// TIA Portal V19 export
FUNCTION_BLOCK "TIMER"   // FB5, LAD
{ S7_Optimized_Access := 'TRUE' }
// stored: MemoryReserve 100, SetENOAutomatically false
   VAR_INPUT
      START_TIMER : Bool;
      HR_SET : Int;
      MIN_SET : Int;
      SEC_SET : Int;
      RESET_TIMER : Bool;
   END_VAR
   VAR_OUTPUT
      SEC : Int;
      MIN : Int;
      HR : Int;
      TIMER_DONE { ExternalAccessible := 'False'; ExternalVisible := 'False'; ExternalWritable := 'False'} : Bool;
   END_VAR
   VAR
      P_TRIG1 : Bool;
      P_TRIG2 : Bool;
      P_TRIG3 : Bool;
   END_VAR
   VAR_TEMP   // added for the SCL form of the ladder/FBD networks
      _w1 : Bool;
      _w2 : Bool;
      _w3 : Bool;
      _w4 : Bool;
   END_VAR
BEGIN

REGION Network 1
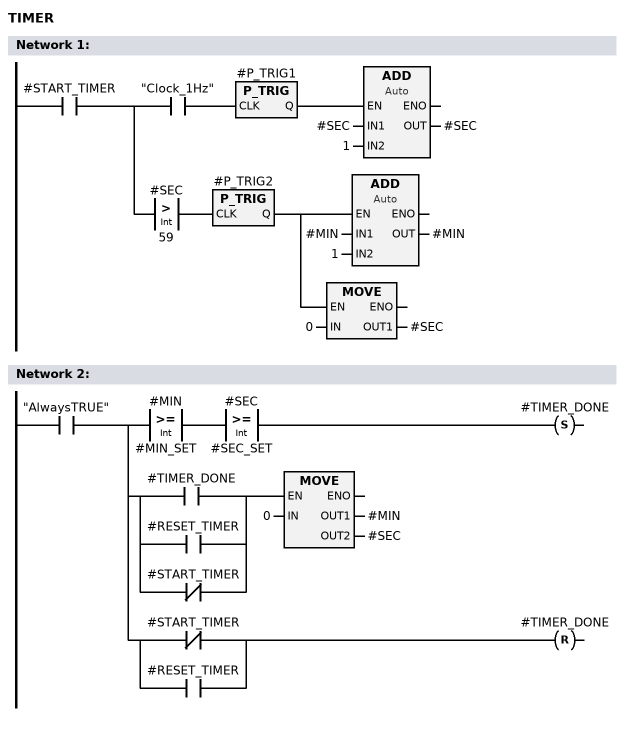
   RUNG wire#powerrail
      Contact( #START_TIMER )
      wire#w1
      Contact( "Clock_1Hz" )
      P_Trig( #P_TRIG1 )
      Add(in1 := #SEC, in2 := 1, out => #SEC)
   END_RUNG
   RUNG wire#w1
      { S7_Templates := "SrcType := Int" } GT_Contact(in1 := #SEC, in2 := 59)
      P_Trig( #P_TRIG2 )
      wire#w2
      Add(in1 := #MIN, in2 := 1, out => #MIN)
   END_RUNG
   RUNG wire#w2
      Move(in := 0, out1 => #SEC)
   END_RUNG
   // the same network as SCL:
   #_w1 := #START_TIMER AND "Clock_1Hz";
   #_w2 := #_w1 AND NOT #P_TRIG1;   // rising edge
   #P_TRIG1 := #_w1;
   IF #_w2 THEN #SEC := #SEC + 1; END_IF;
   #_w3 := #START_TIMER AND (#SEC > 59);
   #_w4 := #_w3 AND NOT #P_TRIG2;   // rising edge
   #P_TRIG2 := #_w3;
   IF #_w4 THEN
       #MIN := #MIN + 1;
       #SEC := 0;
   END_IF;
END_REGION

REGION Network 2
   RUNG wire#powerrail
      Contact( "AlwaysTRUE" )
      wire#w1
      { S7_Templates := "SrcType := Int" } GE_Contact(in1 := #MIN, in2 := #MIN_SET)
      { S7_Templates := "SrcType := Int" } GE_Contact(in1 := #SEC, in2 := #SEC_SET)
      S_Coil( #TIMER_DONE )
   END_RUNG
   RUNG wire#w1
      Contact( #TIMER_DONE )
      wire#w2
      Move(in := 0, out1 => #MIN, out2 => #SEC)
   END_RUNG
   RUNG wire#w1
      Contact( #RESET_TIMER )
   END_RUNG wire#w2
   RUNG wire#w1
      I_Contact( #START_TIMER )
   END_RUNG wire#w2
   RUNG wire#w1
      I_Contact( #START_TIMER )
      wire#w3
      R_Coil( #TIMER_DONE )
   END_RUNG
   RUNG wire#w1
      Contact( #RESET_TIMER )
   END_RUNG wire#w3
   // the same network as SCL:
   IF "AlwaysTRUE" AND (#MIN >= #MIN_SET) AND (#SEC >= #SEC_SET) THEN #TIMER_DONE := TRUE; END_IF;
   IF "AlwaysTRUE" AND (#TIMER_DONE OR #RESET_TIMER OR NOT #START_TIMER) THEN
       #MIN := 0;
       #SEC := 0;
   END_IF;
   IF "AlwaysTRUE" AND (NOT #START_TIMER OR #RESET_TIMER) THEN #TIMER_DONE := FALSE; END_IF;
END_REGION
END_FUNCTION_BLOCK
